FUNCTION_BLOCK FeedTimesCalc (* Basic Function Block Type *)
  (* Standard: 61499-2 *)
  (* Version 0.0, 10/7/2026, Schneider Electric, Template *)
  PACKAGE SE.Nereda;
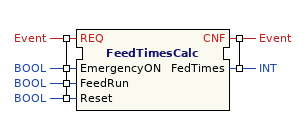
  EVENT_INPUT
    REQ WITH EmergencyON, FeedRun, Reset; (* Normal Execution Request *)
  END_EVENT
  EVENT_OUTPUT
    CNF WITH FedTimes; (* Execution Confirmation *)
  END_EVENT
  VAR_INPUT
    EmergencyON : BOOL; (* Input event qualifier *)
    FeedRun : BOOL;
    Reset : BOOL;
  END_VAR
  VAR_OUTPUT
    FedTimes : INT; (* Output event qualifier *)
  END_VAR
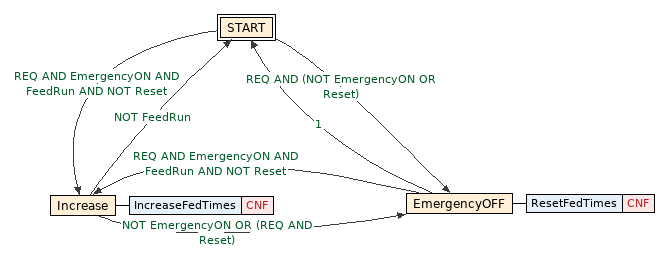
  EC_STATES
    START; (* Initial State *)
    Increase : IncreaseFedTimes -> CNF;
    EmergencyOFF : ResetFedTimes -> CNF;
  END_STATES
  EC_TRANSITIONS
    START TO Increase := REQ AND EmergencyON AND FeedRun AND NOT Reset;
    Increase TO START := NOT FeedRun;
    Increase TO EmergencyOFF := NOT EmergencyON OR (REQ AND Reset);
    START TO EmergencyOFF := REQ AND (NOT EmergencyON OR Reset);
    EmergencyOFF TO START := 1;
    EmergencyOFF TO Increase := REQ AND EmergencyON AND FeedRun AND NOT Reset;
  END_TRANSITIONS
  ALGORITHM IncreaseFedTimes IN ST:
;
FedTimes := FedTimes + 1;
  END_ALGORITHM
  ALGORITHM ResetFedTimes IN ST:
;
FedTimes := 0;
  END_ALGORITHM
END_FUNCTION_BLOCK
